// Minimal I_Focus for the MQTT handler tests: Position is stored by FB_BaseAxis, nothing moves (BROTLib#74).
FUNCTION_BLOCK FB_FocusStub EXTENDS BROTLib.FB_BaseAxis IMPLEMENTS BROTLib.I_Focus
VAR_INPUT
	fMinPosition	: LREAL := -1.0E6;	// travel, as the real focus blocks report it (MONETcommon#122)
	fMaxPosition	: LREAL := 1.0E6;
	nStop			: INT;				// number of Stop() calls
END_VAR

PROPERTY MinPosition : LREAL
GET
MinPosition := fMinPosition;
END_GET
END_PROPERTY

PROPERTY MaxPosition : LREAL
GET
MaxPosition := fMaxPosition;
END_GET
END_PROPERTY

METHOD Stop : BOOL
nStop := nStop + 1;
Stop := TRUE;
END_METHOD

METHOD _StartHoming : BOOL
END_METHOD

END_FUNCTION_BLOCK

(* stored: Version 1.1.0.1, ProductVersion 3.1.4024.15
   POU FB_FocusStub: Id {ba5ff146-f04c-4648-979f-d5c065e2dcc0}, SpecialFunc None
   Property MinPosition: Id {dcb05d04-2922-45aa-a8bd-4dfae8859572}
   Get Get: Id {44935ebe-42c3-47ad-bea6-18679e9b9a5b}
   Property MaxPosition: Id {a844c814-16b5-4cff-90eb-f549351e2ff5}
   Get Get: Id {6e6976cc-dc86-48e9-b887-875be9fa2791}
   Method Stop: Id {0a0dd558-c6f5-49f1-aab9-65d0aa61c69b}
   Method _StartHoming: Id {cff36c3c-f927-4b62-9082-dbd69acf4694} *)
